(* PLC project Unnamed, Unknown Unnamed 1 *)
(* stored: creationDateTime 2026-09-21T13:51:32, modificationDateTime 2026-11-03T16:54:12 *)

PROGRAM waterboiler
  VAR
    STOPPED_STATE : BOOL;
    RUN_STATE : BOOL;
    E_STATE : BOOL;
  END_VAR
  VAR
    START_BTN AT %IX0.0 : BOOL;
    STOP_BTN AT %IX0.1 : BOOL;
    E_STOP AT %IX0.2 : BOOL;
    TEMP_UP AT %IX0.3 : BOOL;
    TEMP_DWN AT %IX0.4 : BOOL;
    P_SWITCH AT %IX0.5 : BOOL;
    HEATER AT %QX0.0 : BOOL;
    LED0 AT %QX0.1 : BOOL;
    LED1 AT %QX0.2 : BOOL;
    LED2 AT %QX0.3 : BOOL;
    LED3 AT %QX0.4 : BOOL;
    LED4 AT %QX0.5 : BOOL;
    LED5 AT %QX0.6 : BOOL;
    E_LED AT %QX0.7 : BOOL;
    SETPOINT AT %MW0 : INT := 80;  (* Default temperature. Min = 80C. Address 32 *)
  END_VAR
  VAR
    POWER : REAL;  (* Represents heating power output *)
  END_VAR
  VAR
    ACTUAL_TEMPERATURE AT %MW1 : INT;
    DIAL_VALUE AT %IW0 : INT;  (* Temp dial = simulates actual temperature *)
  END_VAR
  VAR
    SR0 : SR;
    R_TRIG0 : R_TRIG;
    R_TRIG1 : R_TRIG;
    CTUD0 : CTUD;
    PWM_CONTROLLER0 : PWM_CONTROLLER;
    SERVO_OK : BOOL;
  END_VAR
  VAR
    ANGLE AT %QW0.1 : INT;  (* to test update the servo angle 37 *)
  END_VAR
  VAR
    DUTY : REAL;
    dial_voltage : REAL;  (* actual power usage value *)
    R_TRIG2 : R_TRIG;
    PID0 : PID;
  END_VAR
  VAR  (* added by the conversion: wires and edge detectors of the diagram *)
    _LT198_ENO : BOOL;
    _LT198_OUT : BOOL;
    R_TRIG1_2 : R_TRIG;
    R_TRIG2_2 : R_TRIG;
    _EQ22_OUT : BOOL;
    _EQ23_OUT : BOOL;
    _EQ33_OUT : BOOL;
    _EQ42_OUT : BOOL;
    _EQ50_OUT : BOOL;
    _DIV120_ENO : BOOL;
    _DIV120_OUT : REAL;
    _MUL121_OUT : REAL;
    _GT259_ENO : BOOL;
    _GT259_OUT : BOOL;
  END_VAR

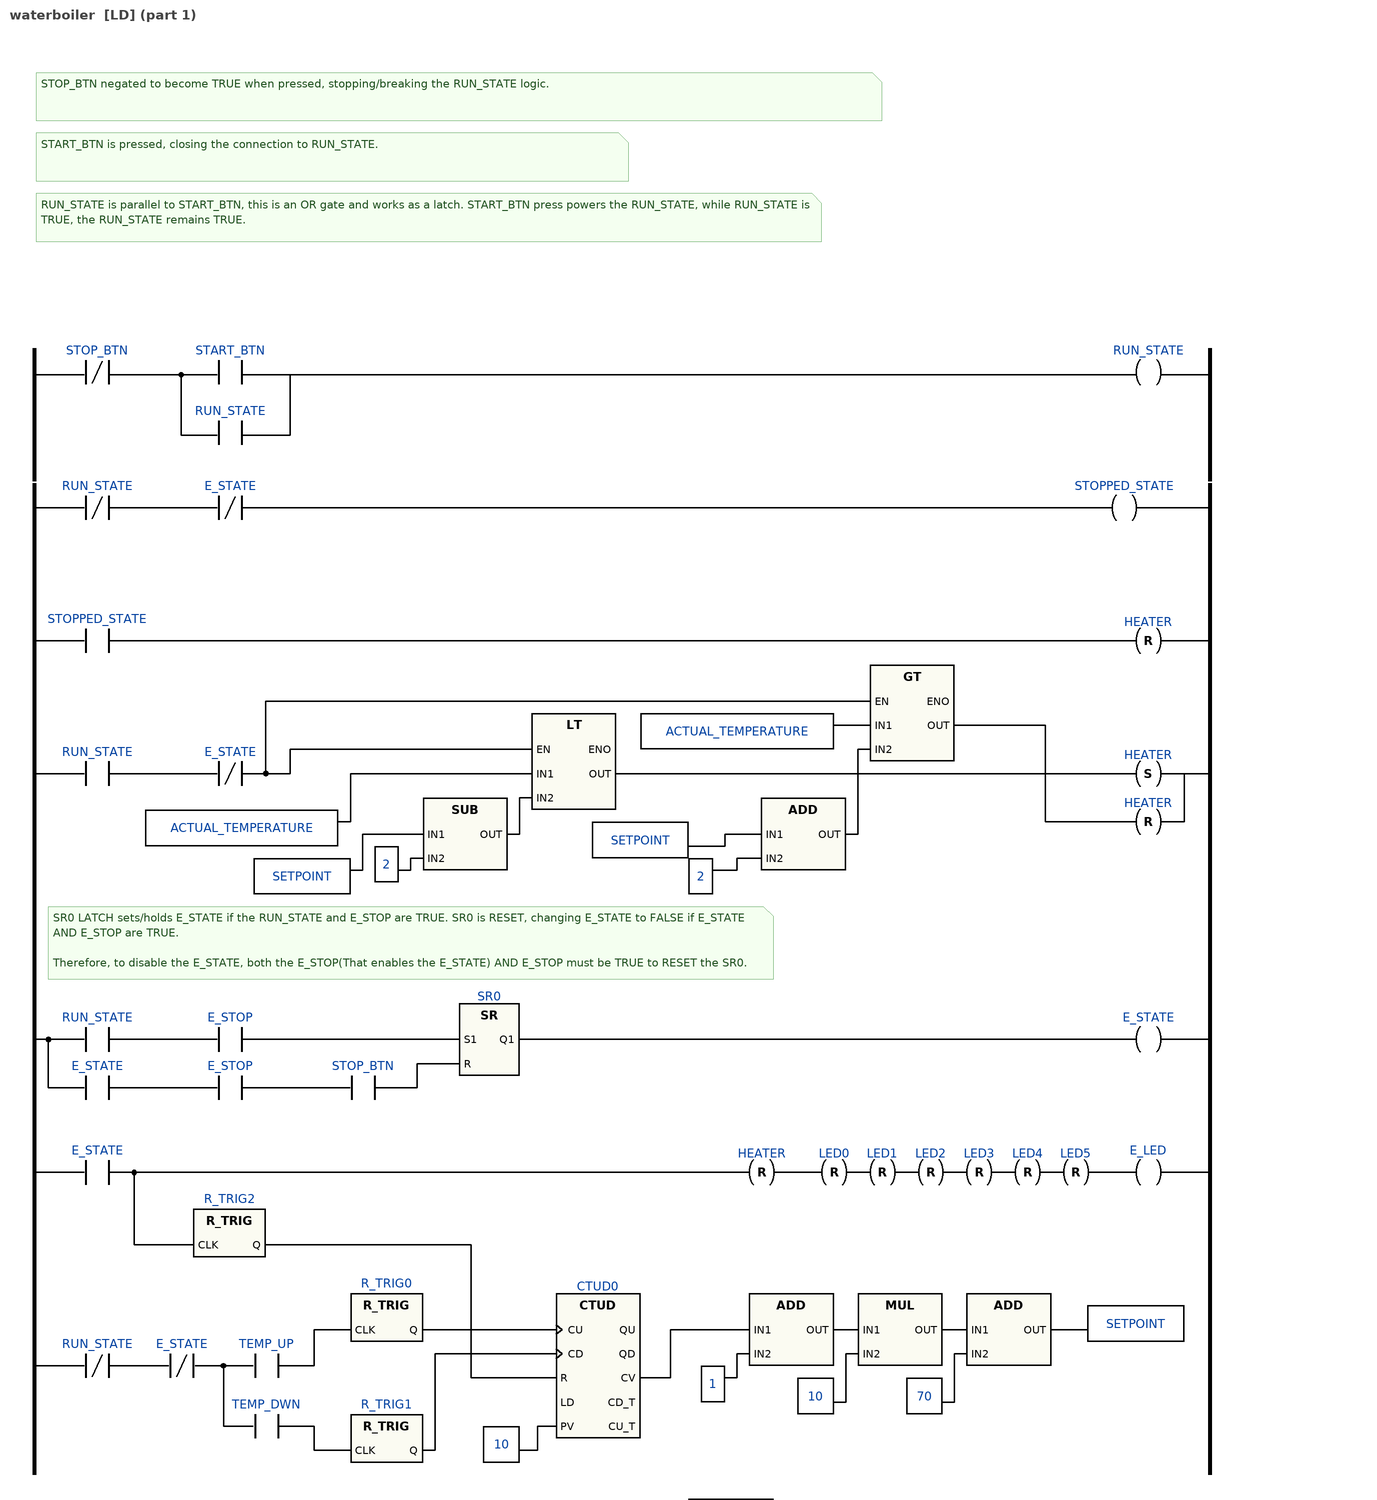
(* LD diagram, written out as Structured Text *)
(* STOP_BTN negated to become TRUE when pressed, stopping/breaking the RUN_STATE logic. *)
(* START_BTN is pressed, closing the connection to RUN_STATE. *)
(* RUN_STATE is parallel to START_BTN, this is an OR gate and works as a latch. START_BTN press powers the RUN_STATE, while RUN_STATE is TRUE, the RUN_STATE remains TRUE. *)
RUN_STATE := NOT STOP_BTN AND (START_BTN OR RUN_STATE);
STOPPED_STATE := NOT RUN_STATE AND NOT E_STATE;
_LT198_OUT := LT(EN := RUN_STATE AND NOT E_STATE, IN1 := ACTUAL_TEMPERATURE, IN2 := SETPOINT - 2, ENO => _LT198_ENO);
IF _LT198_OUT THEN HEATER := TRUE; END_IF;
(* SR0 LATCH sets/holds E_STATE if the RUN_STATE and E_STOP are TRUE. SR0 is RESET, changing E_STATE to FALSE if E_STATE AND E_STOP are TRUE.

Therefore, to disable the E_STATE, both the E_STOP(That enables the E_STATE) AND E_STOP must be TRUE to RESET the SR0. *)
SR0(S1 := RUN_STATE AND E_STOP, R := E_STATE AND E_STOP AND STOP_BTN);
E_STATE := SR0.Q1;
E_LED := E_STATE;
R_TRIG0(CLK := NOT RUN_STATE AND NOT E_STATE AND TEMP_UP);
R_TRIG1_2(CLK := R_TRIG0.Q);
R_TRIG1(CLK := NOT RUN_STATE AND NOT E_STATE AND TEMP_DWN);
R_TRIG2_2(CLK := R_TRIG1.Q);
R_TRIG2(CLK := E_STATE);
CTUD0(CU := R_TRIG1_2.Q, CD := R_TRIG2_2.Q, R := R_TRIG2.Q, PV := 10);
SETPOINT := (CTUD0.CV + 1) * 10 + 70;
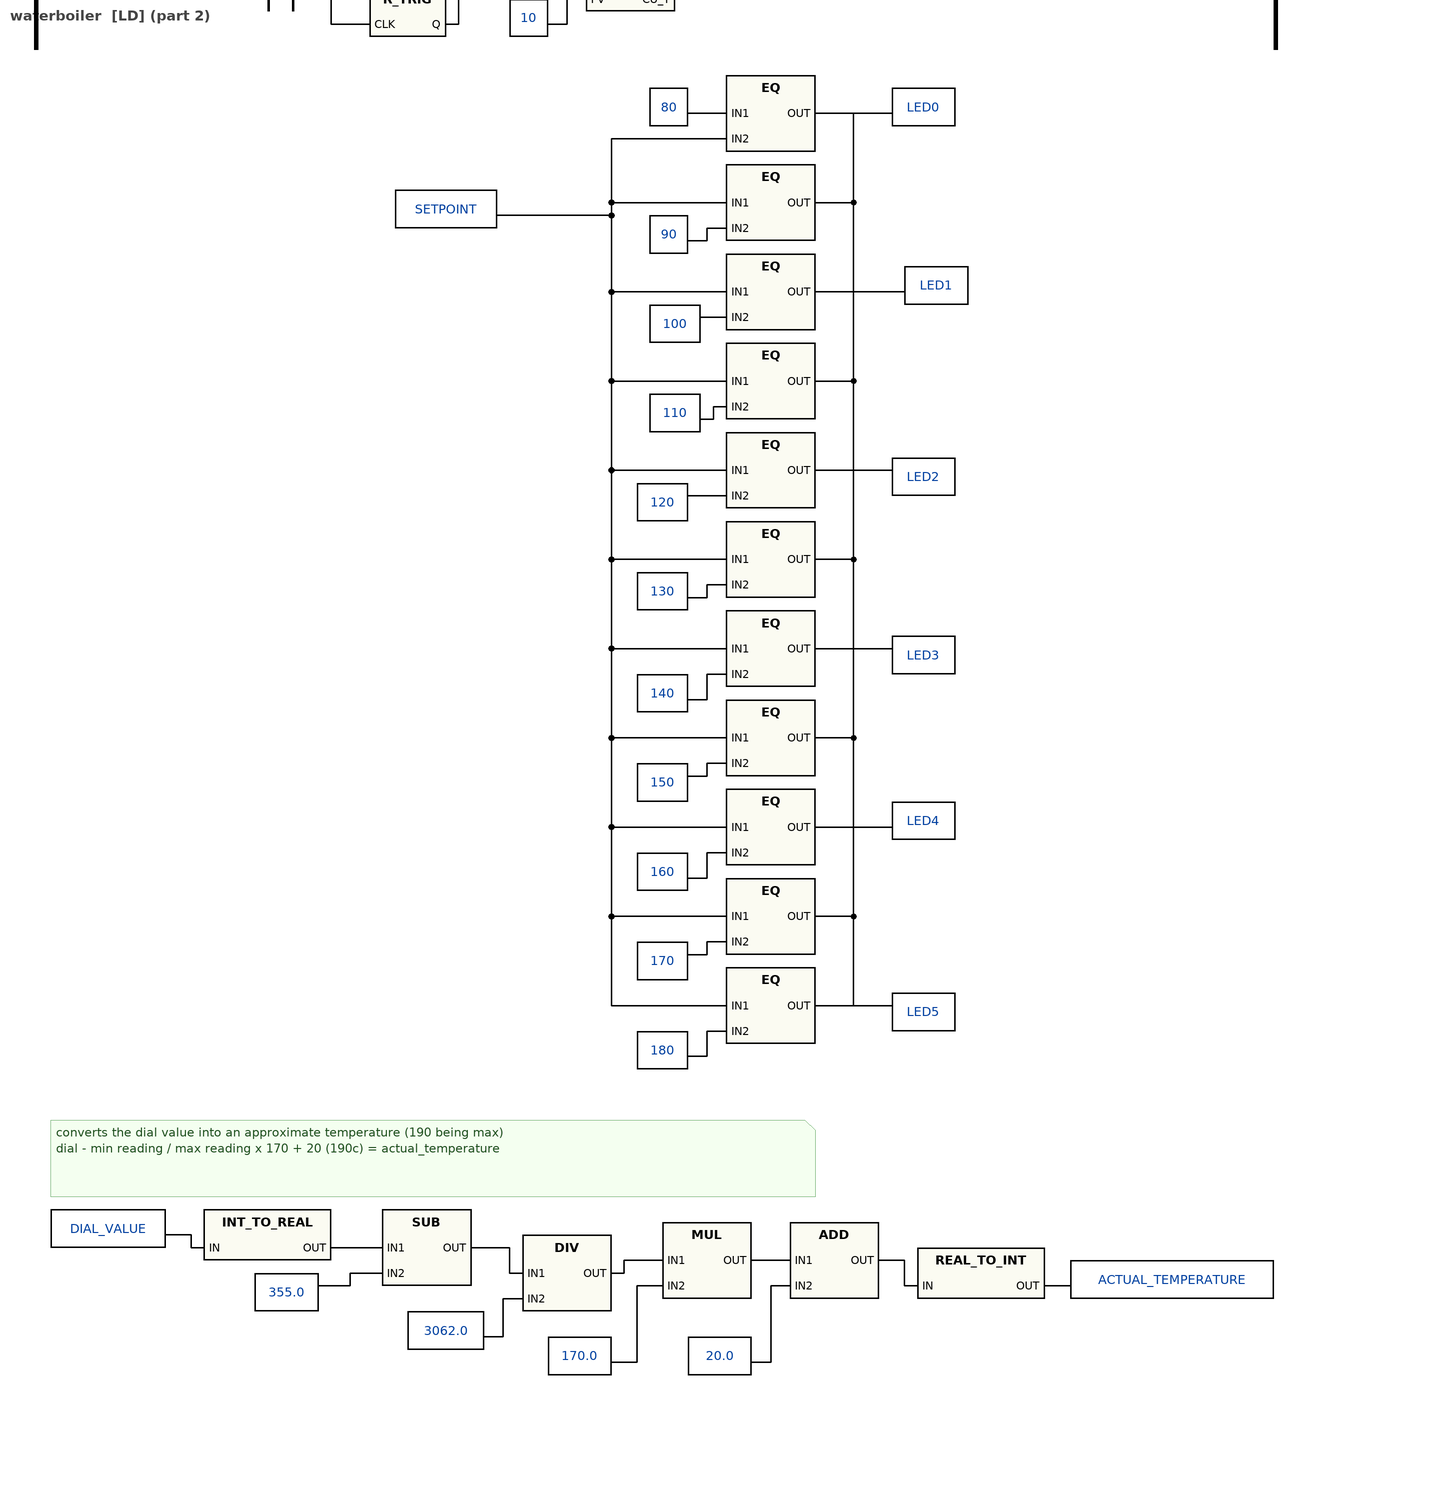
_EQ22_OUT := SETPOINT = 90;
LED0 := 80 = SETPOINT OR _EQ22_OUT;
_EQ23_OUT := SETPOINT = 110;
LED1 := SETPOINT = 100 OR _EQ22_OUT OR _EQ23_OUT;
_EQ33_OUT := SETPOINT = 130;
LED2 := SETPOINT = 120 OR _EQ23_OUT OR _EQ33_OUT;
_EQ42_OUT := SETPOINT = 150;
LED3 := SETPOINT = 140 OR _EQ33_OUT OR _EQ42_OUT;
_EQ50_OUT := SETPOINT = 170;
LED4 := SETPOINT = 160 OR _EQ42_OUT OR _EQ50_OUT;
LED5 := SETPOINT = 180 OR _EQ50_OUT;
IF E_STATE THEN LED0 := FALSE; END_IF;
IF E_STATE THEN LED1 := FALSE; END_IF;
IF E_STATE THEN LED2 := FALSE; END_IF;
IF E_STATE THEN LED3 := FALSE; END_IF;
IF E_STATE THEN LED4 := FALSE; END_IF;
IF E_STATE THEN LED5 := FALSE; END_IF;
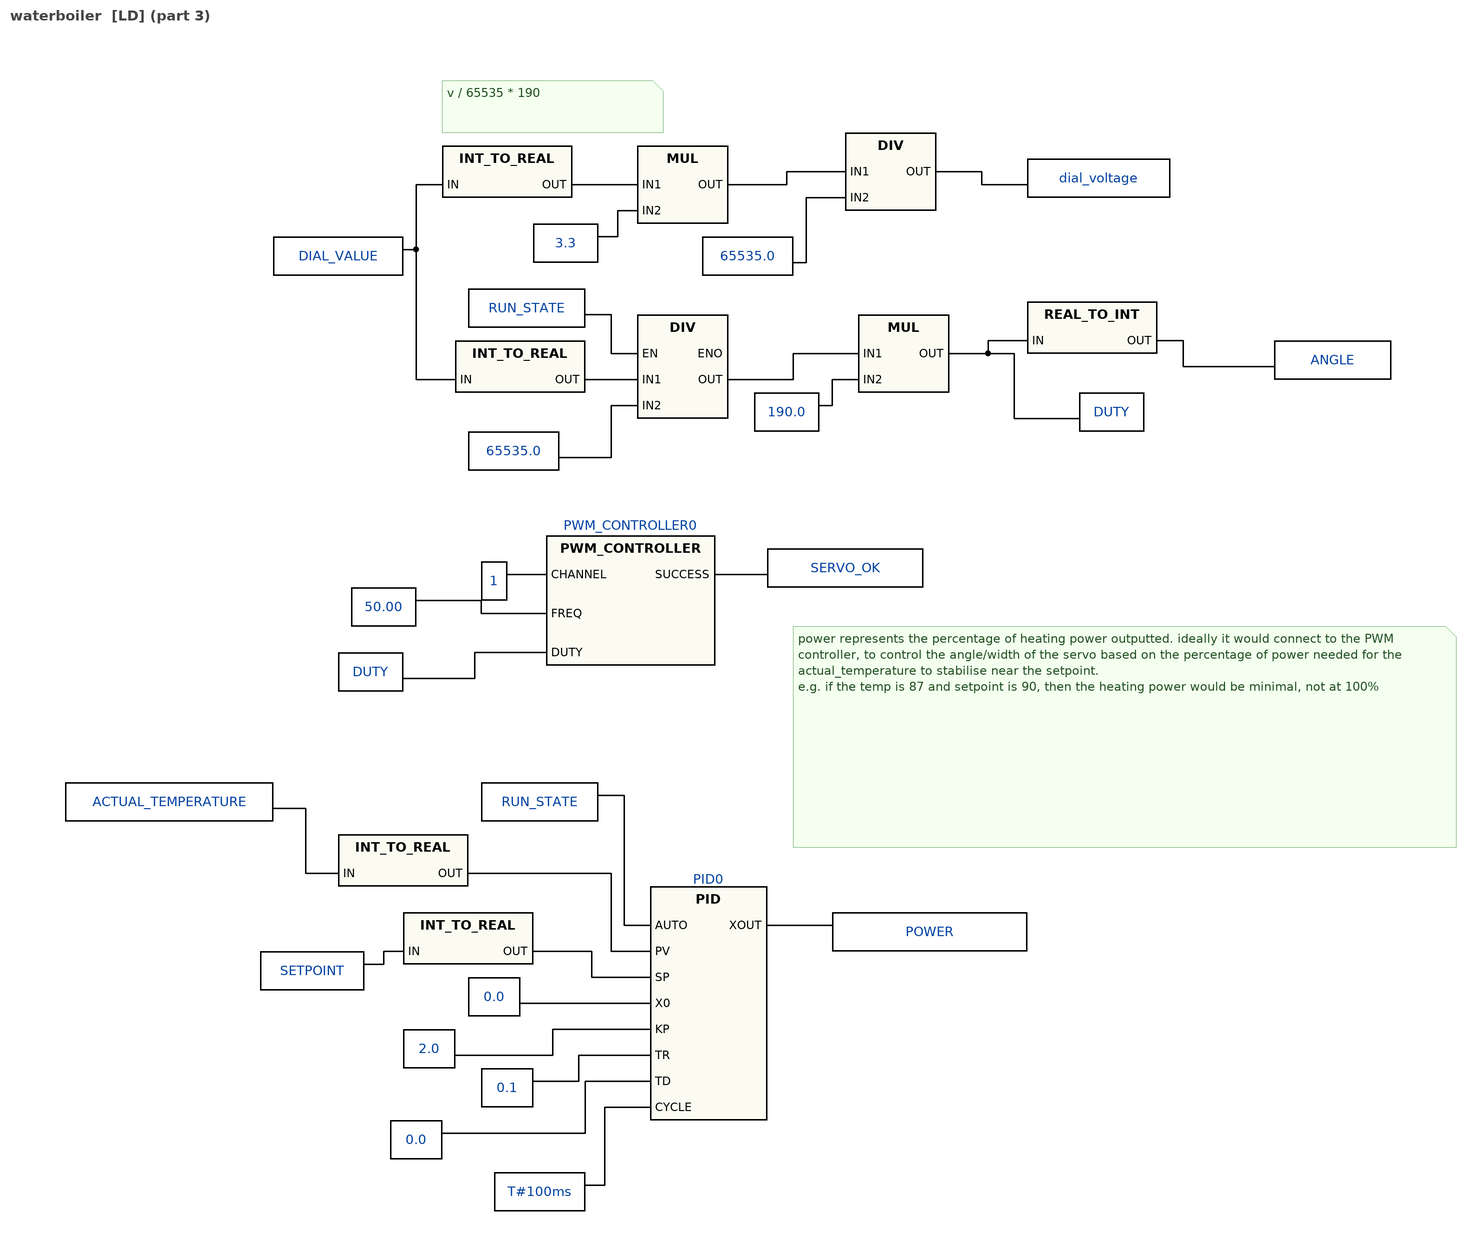
(* converts the dial value into an approximate temperature (190 being max)
dial - min reading / max reading x 170 + 20 (190c) = actual_temperature *)
(* v / 65535 * 190 *)
PWM_CONTROLLER0(CHANNEL := 1, FREQ := 50.00, DUTY := DUTY);
SERVO_OK := PWM_CONTROLLER0.SUCCESS;
_DIV120_OUT := DIV(EN := RUN_STATE, IN1 := INT_TO_REAL(DIAL_VALUE), IN2 := 65535.0, ENO => _DIV120_ENO);
_MUL121_OUT := _DIV120_OUT * 190.0;
DUTY := _MUL121_OUT;
ACTUAL_TEMPERATURE := REAL_TO_INT((INT_TO_REAL(DIAL_VALUE) - 355.0) / 3062.0 * 170.0 + 20.0);
(* power represents the percentage of heating power outputted. ideally it would connect to the PWM controller, to control the angle/width of the servo based on the percentage of power needed for the actual_temperature to stabilise near the setpoint.
e.g. if the temp is 87 and setpoint is 90, then the heating power would be minimal, not at 100% *)
PID0(AUTO := RUN_STATE, PV := INT_TO_REAL(ACTUAL_TEMPERATURE), SP := INT_TO_REAL(SETPOINT), X0 := 0.0, KP := 2.0, TR := 0.1, TD := 0.0, CYCLE := T#100ms);
POWER := PID0.XOUT;
dial_voltage := INT_TO_REAL(DIAL_VALUE) * 3.3 / 65535.0;
ANGLE := REAL_TO_INT(_MUL121_OUT);
_GT259_OUT := GT(EN := RUN_STATE AND NOT E_STATE, IN1 := ACTUAL_TEMPERATURE, IN2 := SETPOINT + 2, ENO => _GT259_ENO);
IF _GT259_OUT THEN HEATER := FALSE; END_IF;
IF E_STATE THEN HEATER := FALSE; END_IF;
IF STOPPED_STATE THEN HEATER := FALSE; END_IF;
END_PROGRAM

CONFIGURATION Config0
  RESOURCE Res0 ON PLC
    TASK task0(INTERVAL := T#20ms, PRIORITY := 0);
    PROGRAM instance0 WITH task0 : waterboiler;
  END_RESOURCE
END_CONFIGURATION
